Fanuc KAREL source: KX00007.KL

PROGRAM KX00007
%NOLOCKGROUP
VAR
  I: INTEGER
  J: INTEGER
  B: BOOLEAN
  F: FILE
  S: STRING[80]
  P: XYZWPR
BEGIN
  PULSE DOUT[1] FOR 100 NOWAIT
END KX00007
